Staubli VAL3: Lab2A_L3.pjx

--- Lab2A_L3.pjx ---
parameters version=s6.8 stackSize=5000 millimeterUnit=true
program file=start.pgx
program file=pickAndPlace.pgx
program file=stop.pgx
program file=physicalIO.pgx
data file=Lab2A_L3.dtx
alias name=io interface=io autoload=true

--- Lab2A_L3.dtx ---


--- start.pgx ---
program start()
// Lab2A Level 3 - shared manual simulation / physical cycle
  local num rowIndex
  local num columnIndex
  local num targetIndex
  local pointRs targetPose
begin

  // Initial state and execution mode.
  userPage()
  cls()
  physicalRun = !simulation

  cycleStep = 0
  placedCount[0] = 0
  placedCount[1] = 0

  vacuumOn = false
  blowOn = false
  trolleyOn = false
  nonMetalGate = false
  metalGate = false
  barrierClosed = true

  ioReady = false
  // Connect physical I/O only on the real station.
  if physicalRun
    taskCreate "physicalIO", 10, physicalIO()
    wait(ioReady == true)
    putln("Lab2A Level 3 - PHYSICAL MODE")
  else
    putln("Lab2A Level 3 - MANUAL SIMULATION")
  endIf

  moveSpeed.vel = 10
  moveSpeed.accel = 10
  moveSpeed.decel = 10
  moveSpeed.blend = off

  // Build the matrix from two taught references: Y+60 mm, approaches Z+50 mm.
  for rowIndex = 0 to 1
    for columnIndex = 0 to 3
      targetIndex = 4*rowIndex + columnIndex
      targetPose = jointToPoint(vacuumTool, world, placePose[4*rowIndex])
      targetPose.trsf.y = targetPose.trsf.y + 60*columnIndex

      if columnIndex != 0
        if !pointToJoint(vacuumTool, placePose[4*rowIndex], targetPose, placePose[targetIndex])
          putln("ERROR: unreachable matrix destination")
          putln(targetIndex)
          return
        endIf
      endIf

      targetPose.trsf.z = targetPose.trsf.z + 50
      if !pointToJoint(vacuumTool, placePose[targetIndex], targetPose, placeApproach[targetIndex])
        putln("ERROR: unreachable matrix approach")
        putln(targetIndex)
        return
      endIf

    endFor

  endFor

  trolleyOn = true
  movej(homePose, vacuumTool, moveSpeed)
  waitEndMove()

  // Classify and place parts until both material groups contain four.
  while placedCount[0] < 4 or placedCount[1] < 4

    cycleStep = 20
    putln("20 - Set partIsMetal, then partAtClass=true")
    wait(partAtClass == true)

    if partIsMetal
      materialType = 1
    else
      materialType = 0
    endIf

    cycleStep = 30
    putln("30 - Select route; actuator settling delay")
    nonMetalGate = materialType == 0
    metalGate = materialType == 1
    delay(0.5)

    cycleStep = 40
    putln("40 - Barrier pulse; then wait partAtRamp=true")
    barrierClosed = false
    delay(0.4)
    barrierClosed = true
    wait(partAtRamp == true)

    cycleStep = 50
    putln("50 - Wait: partAtRamp=false")
    wait(partAtRamp == false)
    if physicalRun
      delay(0.5)
    endIf

    // Skip pickup when this material already has four placed parts.
    if placedCount[materialType] < 4
      placeIndex = 4*materialType + placedCount[materialType]
      call pickAndPlace()
      placedCount[materialType] = placedCount[materialType] + 1
      cycleStep = 80
      putln("80 - Piece placed; next classification part")
      putln("Non-metal placed:")
      putln(placedCount[0])
      putln("Metal placed:")
      putln(placedCount[1])
    else
      cycleStep = 80
      putln("80 - Row full: part passed without pickup; next part")
    endIf

  endWhile

  trolleyOn = false
  barrierClosed = true
  cycleStep = 100
  putln("100 - Completed: four parts of each material")
end

--- physicalIO.pgx ---
program physicalIO()
// Lab2A Level 3 - shared manual simulation / physical cycle
begin

  while true

    // Read sensors.
    partOnTool  = (io:bIn0 == true)
    partAtClass = (io:bIn1 == true)
    partIsMetal = (io:bIn2 == true)
    partAtRamp  = (io:bIn4 == true)

    // Apply output commands; the barrier uses inverted logic.
    io:bOut0 = vacuumOn
    io:bOut1 = blowOn

    io:bOut2 = trolleyOn
    io:bOut3 = nonMetalGate
    io:bOut4 = metalGate
    io:bOut5 = !barrierClosed

    ioReady = true
    delay(0.01)

  endWhile
end

--- pickAndPlace.pgx ---
program pickAndPlace()
// Lab2A Level 3 - shared manual simulation / physical cycle
begin

  // Pick from the selected ramp.
  vacuumOn = false
  blowOn = false

  movej(pickApproach[materialType], vacuumTool, moveSpeed)
  waitEndMove()

  movel(jointToPoint(vacuumTool, world, pickPose[materialType]), vacuumTool, moveSpeed)
  waitEndMove()

  vacuumOn = true
  cycleStep = 60
  putln("60 - Picking part: waiting for vacuum confirmation (partOnTool=true)")
  wait(partOnTool == true)

  movel(jointToPoint(vacuumTool, world, pickApproach[materialType]), vacuumTool, moveSpeed)
  waitEndMove()

  // Transfer and release at the selected destination.
  movej(placeApproach[placeIndex], vacuumTool, moveSpeed)
  waitEndMove()

  movel(jointToPoint(vacuumTool, world, placePose[placeIndex]), vacuumTool, moveSpeed)
  waitEndMove()

  vacuumOn = false
  blowOn = true
  delay(0.3)
  blowOn = false
  cycleStep = 70
  putln("70 - Releasing part: waiting for release confirmation (partOnTool=false)")
  wait(partOnTool == false)

  // Withdraw and return home.
  movel(jointToPoint(vacuumTool, world, placeApproach[placeIndex]), vacuumTool, moveSpeed)
  waitEndMove()

  movej(homePose, vacuumTool, moveSpeed)
  waitEndMove()

end

--- stop.pgx ---
program stop()
// Lab2A Level 3 - shared manual simulation / physical cycle
begin

  // Stop motion and feeding; preserve suction.
  resetMotion()

  trolleyOn = false
  barrierClosed = true
  blowOn = false

  if physicalRun
    taskKill("physicalIO")
    io:bOut2 = false
    io:bOut1 = false
    io:bOut5 = false
  endIf

  cycleStep = -1
  putln("Application stopped safely.")
  resetMotion()

end
